        bool bMarked
        jointRx jJointRx = {j1=-2.687248, j2=16.117165, j3=122.304638, j4=-0.487867, j5=-66.528565, j6=1.978834}
        pointRx pInter
        paraItem pParaItem
          [0]
            bool bSafePoint
            ifItem iIfItem
              [0]
                bool bANDOR[2]
                num nSigIndex[3]
                num nSigType[3]
                num nValue[3]
            mdesc mMdesc
            num nActionIndex = 1
            num nDelay = 5
            num nMoveType = 5
            num nPercentage
            num nSigValue = 1
        pointRx pPointRx[2] = {x=546.855577, y=25.169852, z=121.450925, rx=6.745985, ry=71.76392, rz=-5.460967, shoulder=lefty, elbow=epositive, wrist=wnegative}
        string sID
      [75]
        bool bMarked
        jointRx jJointRx = {j1=-1.639045, j2=12.402747, j3=111.595585, j4=2.517874, j5=-30.594648, j6=-1.669011}
        pointRx pInter
        paraItem pParaItem
          [0]
            bool bSafePoint
            ifItem iIfItem
              [0]
                bool bANDOR[2]
                num nSigIndex[3]
                num nSigType[3]
                num nValue[3]
            mdesc mMdesc
            num nActionIndex = 10
            num nDelay
            num nMoveType = 4
            num nPercentage
            num nSigValue = 1
        pointRx pPointRx[2] = {x=594.549819, y=30.770866, z=171.45682, rx=-40.410864, ry=94.502866, rz=40.920287, shoulder=lefty, elbow=epositive, wrist=wnegative}
        string sID
      [76]
        bool bMarked
        jointRx jJointRx = {j1=-1.639045, j2=12.402747, j3=111.595585, j4=2.517874, j5=-30.594648, j6=-1.669011}
        pointRx pInter
        paraItem pParaItem
          [0]
            bool bSafePoint
            ifItem iIfItem
              [0]
                bool bANDOR[2]
                num nSigIndex[3]
                num nSigType[3]
                num nValue[3]
            mdesc mMdesc
            num nActionIndex = 8
            num nDelay
            num nMoveType = 3
            num nPercentage
            num nSigValue = 1
        pointRx pPointRx[2] = {x=594.549819, y=30.770866, z=171.45682, rx=-40.410864, ry=94.502866, rz=40.920287, shoulder=lefty, elbow=epositive, wrist=wnegative}
        string sID
      [77]
        bool bMarked
        jointRx jJointRx = {j1=-1.639134, j2=22.193742, j3=116.03978, j4=1.817031, j5=-44.819098, j6=-0.790246}
        pointRx pInter
        paraItem pParaItem
          [0]
            bool bSafePoint
            ifItem iIfItem
              [0]
                bool bANDOR[2]
                num nSigIndex[3]
                num nSigType[3]
                num nValue[3]
            mdesc mMdesc = {accel=25, vel=50, leave=1}
            num nActionIndex = 8
            num nDelay = 1.4
            num nMoveType = 7
            num nPercentage
            num nSigValue = 1
        pointRx pPointRx[2] = {x=594.549757, y=30.770873, z=70.540177, rx=-40.399083, ry=94.503271, rz=40.908669, shoulder=lefty, elbow=epositive, wrist=wnegative}
        string sID
      [78]
        bool bMarked
        jointRx jJointRx = {j1=-1.639045, j2=12.402747, j3=111.595585, j4=2.517874, j5=-30.594648, j6=-1.669011}
        pointRx pInter
        paraItem pParaItem
          [0]
            bool bSafePoint
            ifItem iIfItem
              [0]
                bool bANDOR[2]
                num nSigIndex[3]
                num nSigType[3]
                num nValue[3]
            mdesc mMdesc
            num nActionIndex = 10
            num nDelay = 5
            num nMoveType = 4
            num nPercentage
            num nSigValue
        pointRx pPointRx[2] = {x=594.549819, y=30.770866, z=171.45682, rx=-40.410864, ry=94.502866, rz=40.920287, shoulder=lefty, elbow=epositive, wrist=wnegative}
        string sID
      [79]
        bool bMarked
        jointRx jJointRx = {j1=-1.639045, j2=12.402747, j3=111.595585, j4=2.517874, j5=-30.594648, j6=-1.669011}
        pointRx pInter
        paraItem pParaItem
          [0]
            bool bSafePoint
            ifItem iIfItem
              [0]
                bool bANDOR[2]
                num nSigIndex[3]
                num nSigType[3]
                num nValue[3]
            mdesc mMdesc
            num nActionIndex = 10
            num nDelay = 0.8
            num nMoveType = 7
            num nPercentage
            num nSigValue
        pointRx pPointRx[2] = {x=594.549819, y=30.770866, z=171.45682, rx=-40.410864, ry=94.502866, rz=40.920287, shoulder=lefty, elbow=epositive, wrist=wnegative}
        string sID
      [80]
        bool bMarked
        jointRx jJointRx = {j1=-1.639045, j2=12.402747, j3=111.595585, j4=2.517874, j5=-30.594648, j6=-1.669011}
        pointRx pInter
        paraItem pParaItem
          [0]
            bool bSafePoint
            ifItem iIfItem
              [0]
                bool bANDOR[2]
                num nSigIndex[3]
                num nSigType[3]
                num nValue[3]
            mdesc mMdesc
            num nActionIndex = 9
            num nDelay = 5
            num nMoveType = 3
            num nPercentage
            num nSigValue = 1
        pointRx pPointRx[2] = {x=594.549819, y=30.770866, z=171.45682, rx=-40.410864, ry=94.502866, rz=40.920287, shoulder=lefty, elbow=epositive, wrist=wnegative}
        string sID
      [81]
        bool bMarked
        jointRx jJointRx = {j1=-1.639045, j2=12.402747, j3=111.595585, j4=2.517874, j5=-30.594648, j6=-1.669011}
        pointRx pInter
        paraItem pParaItem
          [0]
            bool bSafePoint
            ifItem iIfItem
              [0]
                bool bANDOR[2]
                num nSigIndex[3]
                num nSigType[3]
                num nValue[3]
            mdesc mMdesc
            num nActionIndex = 1
            num nDelay = 5
            num nMoveType = 6
            num nPercentage
            num nSigValue
        pointRx pPointRx[2] = {x=594.549819, y=30.770866, z=171.45682, rx=-40.410864, ry=94.502866, rz=40.920287, shoulder=lefty, elbow=epositive, wrist=wnegative}
        string sID
      [82]
        bool bMarked
        jointRx jJointRx = {j1=-1.639045, j2=12.402747, j3=111.595585, j4=2.517874, j5=-30.594648, j6=-1.669011}
        pointRx pInter
        paraItem pParaItem
          [0]
            bool bSafePoint
            ifItem iIfItem
              [0]
                bool bANDOR[2]
                num nSigIndex[3]
                num nSigType[3]
                num nValue[3]
            mdesc mMdesc
            num nActionIndex = 1
            num nDelay = 5
            num nMoveType = 5
            num nPercentage
            num nSigValue
        pointRx pPointRx[2] = {x=594.549819, y=30.770866, z=171.45682, rx=-40.410864, ry=94.502866, rz=40.920287, shoulder=lefty, elbow=epositive, wrist=wnegative}
        string sID
      [83]
        bool bMarked
        jointRx jJointRx = {j1=-6.64534, j2=-3.725729, j3=129.0442629, j4=-6.345717, j5=-34.650341, j6=4.797577}
        pointRx pInter
        paraItem pParaItem
          [0]
            bool bSafePoint
            ifItem iIfItem
              [0]
                bool bANDOR[2]
                num nSigIndex[3]
                num nSigType[3]
                num nValue[3]
            mdesc mMdesc
            num nActionIndex = 1
            num nDelay = 5
            num nMoveType
            num nPercentage
            num nSigValue
        pointRx pPointRx[2] = {x=472.316864, y=1.637201, z=176.949671, rx=-74.711946, ry=93.153371, rz=74.356802, shoulder=lefty, elbow=epositive, wrist=wnegative}
        string sID
      [84]
        bool bMarked
        jointRx jJointRx = {j1=-1.639045, j2=12.402747, j3=111.595585, j4=2.517874, j5=-30.594648, j6=-1.669011}
        pointRx pInter
        paraItem pParaItem
          [0]
            bool bSafePoint
            ifItem iIfItem
              [0]
                bool bANDOR[2]
                num nSigIndex[3]
                num nSigType[3]
                num nValue[3]
            mdesc mMdesc
            num nActionIndex = 11
            num nDelay = 5
            num nMoveType = 4
            num nPercentage
            num nSigValue = 1
        pointRx pPointRx[2] = {x=594.549819, y=30.770866, z=171.45682, rx=-40.410864, ry=94.502866, rz=40.920287, shoulder=lefty, elbow=epositive, wrist=wnegative}
        string sID
      [85]
        bool bMarked
        jointRx jJointRx = {j1=-1.639045, j2=12.402747, j3=111.595585, j4=2.517874, j5=-30.594648, j6=-1.669011}
        pointRx pInter
        paraItem pParaItem
          [0]
            bool bSafePoint
            ifItem iIfItem
              [0]
                bool bANDOR[2]
                num nSigIndex[3]
                num nSigType[3]
                num nValue[3]
            mdesc mMdesc
            num nActionIndex = 10
            num nDelay = 5
            num nMoveType = 3
            num nPercentage
            num nSigValue
        pointRx pPointRx[2] = {x=594.549819, y=30.770866, z=171.45682, rx=-40.410864, ry=94.502866, rz=40.920287, shoulder=lefty, elbow=epositive, wrist=wnegative}
        string sID
      [86]
        bool bMarked
        jointRx jJointRx = {j1=-1.639045, j2=12.402747, j3=111.595585, j4=2.517874, j5=-30.594648, j6=-1.669011}
        pointRx pInter
        paraItem pParaItem
          [0]
            bool bSafePoint
            ifItem iIfItem
              [0]
                bool bANDOR[2]
                num nSigIndex[3]
                num nSigType[3]
                num nValue[3]
            mdesc mMdesc
            num nActionIndex = 9
            num nDelay = 5
            num nMoveType = 4
            num nPercentage
            num nSigValue
        pointRx pPointRx[2] = {x=594.549819, y=30.770866, z=171.45682, rx=-40.410864, ry=94.502866, rz=40.920287, shoulder=lefty, elbow=epositive, wrist=wnegative}
        string sID
      [87]
        bool bMarked
        jointRx jJointRx = {j1=-1.639045, j2=12.402747, j3=111.595585, j4=2.517874, j5=-30.594648, j6=-1.669011}
        pointRx pInter
        paraItem pParaItem
          [0]
            bool bSafePoint
            ifItem iIfItem
              [0]
                bool bANDOR[2]
                num nSigIndex[3]
                num nSigType[3]
                num nValue[3]
            mdesc mMdesc
            num nActionIndex = 11
            num nDelay = 5
            num nMoveType = 4
            num nPercentage
            num nSigValue
        pointRx pPointRx[2] = {x=594.549819, y=30.770866, z=171.45682, rx=-40.410864, ry=94.502866, rz=40.920287, shoulder=lefty, elbow=epositive, wrist=wnegative}
        string sID
    string sID
  [06 nsk bao]
    num nFrameIndex
    num nMoveID
    num nToolIndex
    pointItem pPointItem[76]
      [0]
        bool bMarked
        jointRx jJointRx = {j1=-2.594987, j2=-12.391258, j3=136.392534, j4=0.644488, j5=-30.575639, j6=-0.113504}
        pointRx pInter
        paraItem pParaItem
          [0]
            bool bSafePoint
            ifItem iIfItem
              [0]
                bool bANDOR[2]
                num nSigIndex[3]
                num nSigType[3]
                num nValue[3]
            mdesc mMdesc
            num nActionIndex = 11
            num nDelay
            num nMoveType = 4
            num nPercentage
            num nSigValue
        pointRx pPointRx[2] = {x=412.772469, y=30.77087, z=171.456836, rx=-40.418431, ry=94.503508, rz=40.927655, shoulder=lefty, elbow=epositive, wrist=wnegative}
        string sID
      [1]
        bool bMarked
        jointRx jJointRx = {j1=-2.594987, j2=-12.391258, j3=136.392534, j4=0.644488, j5=-30.575639, j6=-0.113504}
        pointRx pInter
        paraItem pParaItem
          [0]
            bool bSafePoint
            ifItem iIfItem
              [0]
                bool bANDOR[2]
                num nSigIndex[3]
                num nSigType[3]
                num nValue[3]
            mdesc mMdesc
            num nActionIndex = 9
            num nDelay
            num nMoveType = 4
            num nPercentage
            num nSigValue = 1
        pointRx pPointRx[2] = {x=412.772469, y=30.77087, z=171.456836, rx=-40.418431, ry=94.503508, rz=40.927655, shoulder=lefty, elbow=epositive, wrist=wnegative}
        string sID
      [2]
        bool bMarked
        jointRx jJointRx = {j1=-6.648888, j2=-3.725245, j3=129.0447888, j4=-6.34617, j5=-34.648619, j6=4.79455}
        pointRx pInter
        paraItem pParaItem
          [0]
            bool bSafePoint
            ifItem iIfItem
              [0]
                bool bANDOR[2]
                num nSigIndex[3]
                num nSigType[3]
                num nValue[3]
            mdesc mMdesc
            num nActionIndex
            num nDelay
            num nMoveType
            num nPercentage
            num nSigValue
        pointRx pPointRx[2] = {x=472.316162, y=1.608216, z=176.938999, rx=-74.680314, ry=93.157419, rz=74.321932, shoulder=lefty, elbow=epositive, wrist=wnegative}
        string sID
      [3]
        bool bMarked
        jointRx jJointRx = {j1=-13.0416915, j2=13.589121, j3=123.114063, j4=-3.529204, j5=-45.906395, j6=-89.274538}
        pointRx pInter
        paraItem pParaItem
          [0]
            bool bSafePoint
            ifItem iIfItem
              [0]
                bool bANDOR[2]
                num nSigIndex[3]
                num nSigType[3]
                num nValue[3]
            mdesc mMdesc
            num nActionIndex
            num nDelay
            num nMoveType
            num nPercentage
            num nSigValue
        pointRx pPointRx[2] = {x=539.524688, y=-69.110705, z=102.298754, rx=-85.347202, ry=100.541464, rz=-6.268852, shoulder=lefty, elbow=epositive, wrist=wnegative}
        string sID
      [4]
        bool bMarked
        jointRx jJointRx = {j1=-1.639045, j2=12.402747, j3=111.595585, j4=2.517874, j5=-30.594648, j6=-1.669011}
        pointRx pInter
        paraItem pParaItem
          [0]
            bool bSafePoint
            ifItem iIfItem
              [0]
                bool bANDOR[2]
                num nSigIndex[3]
                num nSigType[3]
                num nValue[3]
            mdesc mMdesc
            num nActionIndex = 1
            num nDelay
            num nMoveType = 6
            num nPercentage
            num nSigValue = 1
        pointRx pPointRx[2] = {x=594.549819, y=30.770866, z=171.45682, rx=-40.410864, ry=94.502866, rz=40.920287, shoulder=lefty, elbow=epositive, wrist=wnegative}
        string sID
      [5]
        bool bMarked
        jointRx jJointRx = {j1=-1.639045, j2=12.402747, j3=111.595585, j4=2.517874, j5=-30.594648, j6=-1.669011}
        pointRx pInter
        paraItem pParaItem
          [0]
            bool bSafePoint
            ifItem iIfItem
              [0]
                bool bANDOR[2]
                num nSigIndex[3]
                num nSigType[3]
                num nValue[3]
            mdesc mMdesc
            num nActionIndex = 1
            num nDelay
            num nMoveType = 5
            num nPercentage
            num nSigValue = 1
        pointRx pPointRx[2] = {x=594.549819, y=30.770866, z=171.45682, rx=-40.410864, ry=94.502866, rz=40.920287, shoulder=lefty, elbow=epositive, wrist=wnegative}
        string sID
      [6]
        bool bMarked
        jointRx jJointRx = {j1=-1.639045, j2=12.402747, j3=111.595585, j4=2.517874, j5=-30.594648, j6=-1.669011}
        pointRx pInter
        paraItem pParaItem
          [0]
            bool bSafePoint
            ifItem iIfItem
              [0]
                bool bANDOR[2]
                num nSigIndex[3]
                num nSigType[3]
                num nValue[3]
            mdesc mMdesc
            num nActionIndex = 10
            num nDelay
            num nMoveType = 4
            num nPercentage
            num nSigValue = 1
        pointRx pPointRx[2] = {x=594.549819, y=30.770866, z=171.45682, rx=-40.410864, ry=94.502866, rz=40.920287, shoulder=lefty, elbow=epositive, wrist=wnegative}
        string sID
      [7]
        bool bMarked
        jointRx jJointRx = {j1=-1.639045, j2=12.402747, j3=111.595585, j4=2.517874, j5=-30.594648, j6=-1.669011}
        pointRx pInter
        paraItem pParaItem
          [0]
            bool bSafePoint
            ifItem iIfItem
              [0]
                bool bANDOR[2]
                num nSigIndex[3]
                num nSigType[3]
                num nValue[3]
            mdesc mMdesc
            num nActionIndex = 8
            num nDelay
            num nMoveType = 3
            num nPercentage
            num nSigValue = 1
        pointRx pPointRx[2] = {x=594.549819, y=30.770866, z=171.45682, rx=-40.410864, ry=94.502866, rz=40.920287, shoulder=lefty, elbow=epositive, wrist=wnegative}
        string sID
      [8]
        bool bMarked
        jointRx jJointRx = {j1=-1.639045, j2=12.402747, j3=111.595585, j4=2.517874, j5=-30.594648, j6=-1.669011}
        pointRx pInter
        paraItem pParaItem
          [0]
            bool bSafePoint
            ifItem iIfItem
              [0]
                bool bANDOR[2]
                num nSigIndex[3]
                num nSigType[3]
                num nValue[3]
            mdesc mMdesc
            num nActionIndex = 8
            num nDelay = 1.2
            num nMoveType = 7
            num nPercentage
            num nSigValue = 1
        pointRx pPointRx[2] = {x=594.549819, y=30.770866, z=171.45682, rx=-40.410864, ry=94.502866, rz=40.920287, shoulder=lefty, elbow=epositive, wrist=wnegative}
        string sID
      [9]
        bool bMarked
        jointRx jJointRx = {j1=-1.639045, j2=12.402747, j3=111.595585, j4=2.517874, j5=-30.594648, j6=-1.669011}
        pointRx pInter
        paraItem pParaItem
          [0]
            bool bSafePoint
            ifItem iIfItem
              [0]
                bool bANDOR[2]
                num nSigIndex[3]
                num nSigType[3]
                num nValue[3]
            mdesc mMdesc
            num nActionIndex = 10
            num nDelay = 5
            num nMoveType = 4
            num nPercentage
            num nSigValue
        pointRx pPointRx[2] = {x=594.549819, y=30.770866, z=171.45682, rx=-40.410864, ry=94.502866, rz=40.920287, shoulder=lefty, elbow=epositive, wrist=wnegative}
        string sID
      [10]
        bool bMarked
        jointRx jJointRx = {j1=-1.639045, j2=12.402747, j3=111.595585, j4=2.517874, j5=-30.594648, j6=-1.669011}
        pointRx pInter
        paraItem pParaItem
          [0]
            bool bSafePoint
            ifItem iIfItem
              [0]
                bool bANDOR[2]
                num nSigIndex[3]
                num nSigType[3]
                num nValue[3]
            mdesc mMdesc
            num nActionIndex = 9
            num nDelay = 5
            num nMoveType = 3
            num nPercentage
            num nSigValue = 1
        pointRx pPointRx[2] = {x=594.549819, y=30.770866, z=171.45682, rx=-40.410864, ry=94.502866, rz=40.920287, shoulder=lefty, elbow=epositive, wrist=wnegative}
        string sID
      [11]
        bool bMarked
        jointRx jJointRx = {j1=-8.869066, j2=16.474618, j3=119.163151, j4=25.800079, j5=-47.747596, j6=-109.409378}
        pointRx pInter
        paraItem pParaItem
          [0]
            bool bSafePoint
            ifItem iIfItem
              [0]
                bool bANDOR[2]
                num nSigIndex[3]
                num nSigType[3]
                num nValue[3]
            mdesc mMdesc
            num nActionIndex
            num nDelay
            num nMoveType
            num nPercentage
            num nSigValue
        pointRx pPointRx[2] = {x=558.358066, y=-69.127961, z=102.227605, rx=-88.177273, ry=117.676396, rz=-3.304957, shoulder=lefty, elbow=epositive, wrist=wnegative}
        string sID
      [12]
        bool bMarked
        jointRx jJointRx = {j1=-1.639045, j2=12.402747, j3=111.595585, j4=2.517874, j5=-30.594648, j6=-1.669011}
        pointRx pInter
        paraItem pParaItem
          [0]
            bool bSafePoint
            ifItem iIfItem
              [0]
                bool bANDOR[2]
                num nSigIndex[3]
                num nSigType[3]
                num nValue[3]
            mdesc mMdesc
            num nActionIndex = 1
            num nDelay
            num nMoveType = 6
            num nPercentage
            num nSigValue = 1
        pointRx pPointRx[2] = {x=594.549819, y=30.770866, z=171.45682, rx=-40.410864, ry=94.502866, rz=40.920287, shoulder=lefty, elbow=epositive, wrist=wnegative}
        string sID
      [13]
        bool bMarked
        jointRx jJointRx = {j1=-1.639045, j2=12.402747, j3=111.595585, j4=2.517874, j5=-30.594648, j6=-1.669011}
        pointRx pInter
        paraItem pParaItem
          [0]
            bool bSafePoint
            ifItem iIfItem
              [0]
                bool bANDOR[2]
                num nSigIndex[3]
                num nSigType[3]
                num nValue[3]
            mdesc mMdesc
            num nActionIndex = 1
            num nDelay
            num nMoveType = 5
            num nPercentage
            num nSigValue = 1
        pointRx pPointRx[2] = {x=594.549819, y=30.770866, z=171.45682, rx=-40.410864, ry=94.502866, rz=40.920287, shoulder=lefty, elbow=epositive, wrist=wnegative}
        string sID
      [14]
        bool bMarked
        jointRx jJointRx = {j1=-1.639045, j2=12.402747, j3=111.595585, j4=2.517874, j5=-30.594648, j6=-1.669011}
        pointRx pInter
        paraItem pParaItem
          [0]
            bool bSafePoint
            ifItem iIfItem
              [0]
                bool bANDOR[2]
                num nSigIndex[3]
                num nSigType[3]
                num nValue[3]
            mdesc mMdesc
            num nActionIndex = 10
            num nDelay
            num nMoveType = 4
            num nPercentage
            num nSigValue = 1
        pointRx pPointRx[2] = {x=594.549819, y=30.770866, z=171.45682, rx=-40.410864, ry=94.502866, rz=40.920287, shoulder=lefty, elbow=epositive, wrist=wnegative}
        string sID
      [15]
        bool bMarked
        jointRx jJointRx = {j1=-1.639045, j2=12.402747, j3=111.595585, j4=2.517874, j5=-30.594648, j6=-1.669011}
        pointRx pInter
        paraItem pParaItem
          [0]
            bool bSafePoint
            ifItem iIfItem
              [0]
                bool bANDOR[2]
                num nSigIndex[3]
                num nSigType[3]
                num nValue[3]
            mdesc mMdesc
            num nActionIndex = 8
            num nDelay
            num nMoveType = 3
            num nPercentage
            num nSigValue = 1
        pointRx pPointRx[2] = {x=594.549819, y=30.770866, z=171.45682, rx=-40.410864, ry=94.502866, rz=40.920287, shoulder=lefty, elbow=epositive, wrist=wnegative}
        string sID
      [16]
        bool bMarked
        jointRx jJointRx = {j1=-1.639045, j2=12.402747, j3=111.595585, j4=2.517874, j5=-30.594648, j6=-1.669011}
        pointRx pInter
        paraItem pParaItem
          [0]
            bool bSafePoint
            ifItem iIfItem
              [0]
                bool bANDOR[2]
                num nSigIndex[3]
                num nSigType[3]
                num nValue[3]
            mdesc mMdesc
            num nActionIndex = 8
            num nDelay = 1.2
            num nMoveType = 7
            num nPercentage
            num nSigValue = 1
        pointRx pPointRx[2] = {x=594.549819, y=30.770866, z=171.45682, rx=-40.410864, ry=94.502866, rz=40.920287, shoulder=lefty, elbow=epositive, wrist=wnegative}
        string sID
      [17]
        bool bMarked
        jointRx jJointRx = {j1=-1.639045, j2=12.402747, j3=111.595585, j4=2.517874, j5=-30.594648, j6=-1.669011}
        pointRx pInter
        paraItem pParaItem
          [0]
            bool bSafePoint
            ifItem iIfItem
              [0]
                bool bANDOR[2]
                num nSigIndex[3]
                num nSigType[3]
                num nValue[3]
            mdesc mMdesc
            num nActionIndex = 10
            num nDelay = 5
            num nMoveType = 4
            num nPercentage
            num nSigValue
        pointRx pPointRx[2] = {x=594.549819, y=30.770866, z=171.45682, rx=-40.410864, ry=94.502866, rz=40.920287, shoulder=lefty, elbow=epositive, wrist=wnegative}
        string sID
      [18]
        bool bMarked
        jointRx jJointRx = {j1=-1.639045, j2=12.402747, j3=111.595585, j4=2.517874, j5=-30.594648, j6=-1.669011}
        pointRx pInter
        paraItem pParaItem
          [0]
            bool bSafePoint
            ifItem iIfItem
              [0]
                bool bANDOR[2]
                num nSigIndex[3]
                num nSigType[3]
                num nValue[3]
            mdesc mMdesc
            num nActionIndex = 9
            num nDelay = 5
            num nMoveType = 3
            num nPercentage
            num nSigValue = 1
        pointRx pPointRx[2] = {x=594.549819, y=30.770866, z=171.45682, rx=-40.410864, ry=94.502866, rz=40.920287, shoulder=lefty, elbow=epositive, wrist=wnegative}
        string sID
      [19]
        bool bMarked
        jointRx jJointRx = {j1=-12.0973934, j2=29.692013, j3=112.730932, j4=-9.94873, j5=-90.923784, j6=35.953063}
        pointRx pInter
        paraItem pParaItem
          [0]
            bool bSafePoint
            ifItem iIfItem
              [0]
                bool bANDOR[2]
                num nSigIndex[3]
                num nSigType[3]
                num nValue[3]
            mdesc mMdesc
            num nActionIndex
            num nDelay
            num nMoveType
            num nPercentage
            num nSigValue
        pointRx pPointRx[2] = {x=597.610117, y=-59.285719, z=93.706544, rx=-0.690577, ry=52.164123, rz=29.161478, shoulder=lefty, elbow=epositive, wrist=wnegative}
        string sID
      [20]
        bool bMarked
        jointRx jJointRx = {j1=-1.639045, j2=12.402747, j3=111.595585, j4=2.517874, j5=-30.594648, j6=-1.669011}
        pointRx pInter
        paraItem pParaItem
          [0]
            bool bSafePoint
            ifItem iIfItem
              [0]
                bool bANDOR[2]
                num nSigIndex[3]
                num nSigType[3]
                num nValue[3]
            mdesc mMdesc
            num nActionIndex = 1
            num nDelay
            num nMoveType = 6
            num nPercentage
            num nSigValue = 1
        pointRx pPointRx[2] = {x=594.549819, y=30.770866, z=171.45682, rx=-40.410864, ry=94.502866, rz=40.920287, shoulder=lefty, elbow=epositive, wrist=wnegative}
        string sID
      [21]
        bool bMarked
        jointRx jJointRx = {j1=-1.639045, j2=12.402747, j3=111.595585, j4=2.517874, j5=-30.594648, j6=-1.669011}
        pointRx pInter
        paraItem pParaItem
          [0]
            bool bSafePoint
            ifItem iIfItem
              [0]
                bool bANDOR[2]
                num nSigIndex[3]
                num nSigType[3]
                num nValue[3]
            mdesc mMdesc
            num nActionIndex = 1
            num nDelay
            num nMoveType = 5
            num nPercentage
            num nSigValue = 1
        pointRx pPointRx[2] = {x=594.549819, y=30.770866, z=171.45682, rx=-40.410864, ry=94.502866, rz=40.920287, shoulder=lefty, elbow=epositive, wrist=wnegative}
        string sID
      [22]
        bool bMarked
        jointRx jJointRx = {j1=-1.639045, j2=12.402747, j3=111.595585, j4=2.517874, j5=-30.594648, j6=-1.669011}
        pointRx pInter
        paraItem pParaItem
          [0]
            bool bSafePoint
            ifItem iIfItem
              [0]
                bool bANDOR[2]
                num nSigIndex[3]
                num nSigType[3]
                num nValue[3]
            mdesc mMdesc
            num nActionIndex = 10
            num nDelay
            num nMoveType = 4
            num nPercentage
            num nSigValue = 1
        pointRx pPointRx[2] = {x=594.549819, y=30.770866, z=171.45682, rx=-40.410864, ry=94.502866, rz=40.920287, shoulder=lefty, elbow=epositive, wrist=wnegative}
        string sID
      [23]
        bool bMarked
        jointRx jJointRx = {j1=-1.639045, j2=12.402747, j3=111.595585, j4=2.517874, j5=-30.594648, j6=-1.669011}
        pointRx pInter
        paraItem pParaItem
          [0]
            bool bSafePoint
            ifItem iIfItem
              [0]
                bool bANDOR[2]
                num nSigIndex[3]
                num nSigType[3]
                num nValue[3]
            mdesc mMdesc
            num nActionIndex = 8
            num nDelay
            num nMoveType = 3
            num nPercentage
            num nSigValue = 1
        pointRx pPointRx[2] = {x=594.549819, y=30.770866, z=171.45682, rx=-40.410864, ry=94.502866, rz=40.920287, shoulder=lefty, elbow=epositive, wrist=wnegative}
        string sID
      [24]
        bool bMarked
        jointRx jJointRx = {j1=-1.639045, j2=12.402747, j3=111.595585, j4=2.517874, j5=-30.594648, j6=-1.669011}
        pointRx pInter
        paraItem pParaItem
          [0]
            bool bSafePoint
            ifItem iIfItem
              [0]
                bool bANDOR[2]
                num nSigIndex[3]
                num nSigType[3]
                num nValue[3]
            mdesc mMdesc
            num nActionIndex = 8
            num nDelay = 2.2
            num nMoveType = 7
            num nPercentage
            num nSigValue = 1
        pointRx pPointRx[2] = {x=594.549819, y=30.770866, z=171.45682, rx=-40.410864, ry=94.502866, rz=40.920287, shoulder=lefty, elbow=epositive, wrist=wnegative}
        string sID
      [25]
        bool bMarked
        jointRx jJointRx = {j1=-1.639045, j2=12.402747, j3=111.595585, j4=2.517874, j5=-30.594648, j6=-1.669011}
        pointRx pInter
        paraItem pParaItem
          [0]
            bool bSafePoint
            ifItem iIfItem
              [0]
                bool bANDOR[2]
                num nSigIndex[3]
                num nSigType[3]
                num nValue[3]
            mdesc mMdesc
            num nActionIndex = 10
            num nDelay = 5
            num nMoveType = 4
            num nPercentage
            num nSigValue
        pointRx pPointRx[2] = {x=594.549819, y=30.770866, z=171.45682, rx=-40.410864, ry=94.502866, rz=40.920287, shoulder=lefty, elbow=epositive, wrist=wnegative}
        string sID
      [26]
        bool bMarked
        jointRx jJointRx = {j1=-1.639045, j2=12.402747, j3=111.595585, j4=2.517874, j5=-30.594648, j6=-1.669011}
        pointRx pInter
        paraItem pParaItem
          [0]
            bool bSafePoint
            ifItem iIfItem
              [0]
                bool bANDOR[2]
                num nSigIndex[3]
                num nSigType[3]
                num nValue[3]
            mdesc mMdesc
            num nActionIndex = 9
            num nDelay = 5
            num nMoveType = 3
            num nPercentage
            num nSigValue = 1
        pointRx pPointRx[2] = {x=594.549819, y=30.770866, z=171.45682, rx=-40.410864, ry=94.502866, rz=40.920287, shoulder=lefty, elbow=epositive, wrist=wnegative}
        string sID
      [27]
        bool bMarked
        jointRx jJointRx = {j1=-3.658412, j2=-3.554964, j3=108.46581, j4=2.353449, j5=5.810977, j6=-2.88172}
        pointRx pInter
        paraItem pParaItem
          [0]
            bool bSafePoint
            ifItem iIfItem
              [0]
                bool bANDOR[2]
                num nSigIndex[3]
                num nSigType[3]
                num nValue[3]
            mdesc mMdesc
            num nActionIndex
            num nDelay
            num nMoveType
            num nPercentage
            num nSigValue
        pointRx pPointRx[2] = {x=530.0109411, y=16.630735, z=279.44816, rx=-8.921642, ry=110.982384, rz=9.0937081, shoulder=lefty, elbow=epositive, wrist=wpositive}
        string sID
      [28]
        bool bMarked
        jointRx jJointRx = {j1=0.670944, j2=16.912776, j3=64.983738, j4=-22.375541, j5=61.12488, j6=-0.704871}
        pointRx pInter
        paraItem pParaItem
          [0]
            bool bSafePoint
            ifItem iIfItem
              [0]
                bool bANDOR[2]
                num nSigIndex[3]
                num nSigType[3]
                num nValue[3]
            mdesc mMdesc
            num nActionIndex
            num nDelay
            num nMoveType
            num nPercentage
            num nSigValue
        pointRx pPointRx[2] = {x=653.37786, y=24.317879, z=393.168061, rx=-23.985387, ry=143.409914, rz=2.3528, shoulder=lefty, elbow=epositive, wrist=wpositive}
        string sID
      [29]
        bool bMarked
        jointRx jJointRx = {j1=-1.639045, j2=12.402747, j3=111.595585, j4=2.517874, j5=-30.594648, j6=-1.669011}
        pointRx pInter
        paraItem pParaItem
          [0]
            bool bSafePoint
            ifItem iIfItem
              [0]
                bool bANDOR[2]
                num nSigIndex[3]
                num nSigType[3]
                num nValue[3]
            mdesc mMdesc
            num nActionIndex = 1
            num nDelay
            num nMoveType = 6
            num nPercentage
            num nSigValue = 1
        pointRx pPointRx[2] = {x=594.549819, y=30.770866, z=171.45682, rx=-40.410864, ry=94.502866, rz=40.920287, shoulder=lefty, elbow=epositive, wrist=wnegative}
        string sID
      [30]
        bool bMarked
        jointRx jJointRx = {j1=-1.639045, j2=12.402747, j3=111.595585, j4=2.517874, j5=-30.594648, j6=-1.669011}
        pointRx pInter
        paraItem pParaItem
          [0]
            bool bSafePoint
            ifItem iIfItem
              [0]
                bool bANDOR[2]
                num nSigIndex[3]
                num nSigType[3]
                num nValue[3]
            mdesc mMdesc
            num nActionIndex = 1
            num nDelay
            num nMoveType = 5
            num nPercentage
            num nSigValue = 1
        pointRx pPointRx[2] = {x=594.549819, y=30.770866, z=171.45682, rx=-40.410864, ry=94.502866, rz=40.920287, shoulder=lefty, elbow=epositive, wrist=wnegative}
        string sID
      [31]
        bool bMarked
        jointRx jJointRx = {j1=-1.639045, j2=12.402747, j3=111.595585, j4=2.517874, j5=-30.594648, j6=-1.669011}
        pointRx pInter
        paraItem pParaItem
          [0]
            bool bSafePoint
            ifItem iIfItem
              [0]
                bool bANDOR[2]
                num nSigIndex[3]
                num nSigType[3]
                num nValue[3]
            mdesc mMdesc
            num nActionIndex = 10
            num nDelay
            num nMoveType = 4
            num nPercentage
            num nSigValue = 1
        pointRx pPointRx[2] = {x=594.549819, y=30.770866, z=171.45682, rx=-40.410864, ry=94.502866, rz=40.920287, shoulder=lefty, elbow=epositive, wrist=wnegative}
        string sID
      [32]
        bool bMarked
        jointRx jJointRx = {j1=-1.639045, j2=12.402747, j3=111.595585, j4=2.517874, j5=-30.594648, j6=-1.669011}
        pointRx pInter
        paraItem pParaItem
          [0]
            bool bSafePoint
            ifItem iIfItem
